Staubli VAL3: updateStr.pgx

public program updateStr(num x_nItemIn, string& x_sTextOut, string x_sComment)
begin
  switch sLanguage
    case "chinese"
      x_sTextOut=sHmiCN[x_nItemIn]
    break
    //
    case "english"
      x_sTextOut=sHmiEN[x_nItemIn]
    break
  endSwitch
end
